MOVL C00866 V=7.0 ACC=20 DEC=20
MOVL C00867 V=7.0 ACC=20 DEC=20
MOVL C00868 V=7.0 ACC=20 DEC=20
MOVL C00869 V=7.0 ACC=20 DEC=20
MOVL C00870 V=7.0 ACC=20 DEC=20
MOVL C00871 V=7.0 ACC=20 DEC=20
MOVL C00872 V=7.0 ACC=20 DEC=20
MOVL C00873 V=7.0 ACC=20 DEC=20
MOVL C00874 V=7.0 ACC=20 DEC=20
MOVL C00875 V=7.0 ACC=20 DEC=20
MOVL C00876 V=7.0 ACC=20 DEC=20
MOVL C00877 V=7.0 ACC=20 DEC=20
MOVL C00878 V=7.0 PL=1
MOVL C00879 V=7.0 ACC=20 DEC=20
MOVL C00880 V=7.0 ACC=20 DEC=20
MOVL C00881 V=7.0 ACC=20 DEC=20
MOVL C00882 V=7.0 ACC=20 DEC=20
MOVL C00883 V=7.0 ACC=20 DEC=20
MOVL C00884 V=7.0 ACC=20 DEC=20
MOVL C00885 V=7.0 ACC=20 DEC=20
MOVL C00886 V=7.0 ACC=20 DEC=20
MOVL C00887 V=7.0 ACC=20 DEC=20
MOVL C00888 V=11.0 ACC=20 DEC=20
MOVC C00889 V=11.0 ACC=20 DEC=20
MOVC C00890 V=11.0 ACC=20 DEC=20
MOVC C00891 V=11.0 ACC=20 DEC=20
MOVL C00892 V=7.0 ACC=20 DEC=20
MOVL C00893 V=7.0 ACC=20 DEC=20
MOVL C00894 V=7.0 ACC=20 DEC=20
MOVL C00895 V=7.0 ACC=20 DEC=20
MOVL C00896 V=7.0 ACC=20 DEC=20
MOVL C00897 V=7.0 ACC=20 DEC=20
MOVL C00898 V=7.0 ACC=20 DEC=20
MOVL C00899 V=7.0 ACC=20 DEC=20
MOVL C00900 V=7.0 ACC=20 DEC=20
MOVL C00901 V=7.0 ACC=20 DEC=20
MOVL C00902 V=7.0 ACC=20 DEC=20
MOVL C00903 V=7.0 ACC=20 DEC=20
MOVL C00904 V=7.0 ACC=20 DEC=20
MOVL C00905 V=7.0 ACC=20 DEC=20
MOVL C00906 V=7.0 ACC=20 DEC=20
MOVL C00907 V=7.0 ACC=20 DEC=20
MOVL C00908 V=7.0 ACC=20 DEC=20
MOVL C00909 V=7.0 ACC=20 DEC=20
MOVL C00910 V=7.0 ACC=20 DEC=20
MOVL C00911 V=7.0 ACC=20 DEC=20
ARCOF
TIMER T=30.00
MOVL C00912 V=11.0 ACC=20 DEC=20
*LAG11
MACRO1 MJ#(0) ARGF2
ARCON
MOVL C00913 V=7.0 ACC=20 DEC=20
MOVL C00914 V=7.0 ACC=20 DEC=20
MOVL C00915 V=7.0 ACC=20 DEC=20
MOVL C00916 V=7.0 ACC=20 DEC=20
MOVL C00917 V=7.0 ACC=20 DEC=20
MOVL C00918 V=7.0 ACC=20 DEC=20
MOVL C00919 V=7.0 ACC=20 DEC=20
MOVL C00920 V=7.0 ACC=20 DEC=20
MOVL C00921 V=7.0 ACC=20 DEC=20
MOVL C00922 V=7.0 ACC=20 DEC=20
MOVL C00923 V=7.0 ACC=20 DEC=20
MOVL C00924 V=7.0 ACC=20 DEC=20
MOVL C00925 V=7.0 ACC=20 DEC=20
MOVL C00926 V=7.0 ACC=20 DEC=20
MOVL C00927 V=7.0 ACC=20 DEC=20
MOVL C00928 V=7.0 ACC=20 DEC=20
MOVL C00929 V=7.0 ACC=20 DEC=20
MOVL C00930 V=7.0 ACC=20 DEC=20
MOVL C00931 V=7.0 ACC=20 DEC=20
MOVL C00932 V=11.0 ACC=20 DEC=20
MOVC C00933 V=11.0 ACC=20 DEC=20
MOVC C00934 V=11.0 ACC=20 DEC=20
MOVC C00935 V=11.0 ACC=20 DEC=20
MOVL C00936 V=7.0 ACC=20 DEC=20
MOVL C00937 V=7.0 ACC=20 DEC=20
MOVL C00938 V=7.0 ACC=20 DEC=20
MOVL C00939 V=7.0 ACC=20 DEC=20
MOVL C00940 V=7.0 ACC=20 DEC=20
MOVL C00941 V=7.0 ACC=20 DEC=20
MOVL C00942 V=7.0 ACC=20 DEC=20
MOVL C00943 V=7.0 ACC=20 DEC=20
MOVL C00944 V=7.0 ACC=20 DEC=20
MOVL C00945 V=7.0 PL=1
MOVL C00946 V=7.0 ACC=20 DEC=20
MOVL C00947 V=7.0 ACC=20 DEC=20
MOVL C00948 V=7.0 ACC=20 DEC=20
MOVL C00949 V=7.0 ACC=20 DEC=20
MOVL C00950 V=7.0 ACC=20 DEC=20
MOVL C00951 V=7.0 ACC=20 DEC=20
MOVL C00952 V=7.0 ACC=20 DEC=20
MOVL C00953 V=7.0 ACC=20 DEC=20
MOVL C00954 V=7.0 ACC=20 DEC=20
MOVL C00955 V=7.0 ACC=20 DEC=20
MOVL C00956 V=7.0 ACC=20 DEC=20
MOVL C00957 V=7.0 ACC=20 DEC=20
MOVL C00958 V=7.0 ACC=20 DEC=20
MOVL C00959 V=7.0 ACC=20 DEC=20
MOVL C00960 V=7.0 ACC=20 DEC=20
MOVL C00961 V=7.0 ACC=20 DEC=20
MOVL C00962 V=7.0 ACC=20 DEC=20
MOVL C00963 V=7.0 ACC=20 DEC=20
MOVL C00964 V=7.0 ACC=20 DEC=20
MOVL C00965 V=7.0 ACC=20 DEC=20
MOVL C00966 V=7.0 ACC=20 DEC=20
MOVL C00967 V=11.0 ACC=20 DEC=20
MOVC C00968 V=11.0 ACC=20 DEC=20
MOVC C00969 V=11.0 ACC=20 DEC=20
MOVC C00970 V=11.0 ACC=20 DEC=20
MOVL C00971 V=7.0 ACC=20 DEC=20
MOVL C00972 V=7.0 ACC=20 DEC=20
MOVL C00973 V=7.0 ACC=20 DEC=20
MOVL C00974 V=7.0 ACC=20 DEC=20
MOVL C00975 V=7.0 ACC=20 DEC=20
MOVL C00976 V=7.0 ACC=20 DEC=20
MOVL C00977 V=7.0 ACC=20 DEC=20
MOVL C00978 V=7.0 ACC=20 DEC=20
MOVL C00979 V=7.0 ACC=20 DEC=20
MOVL C00980 V=7.0 ACC=20 DEC=20
MOVL C00981 V=7.0 ACC=20 DEC=20
MOVL C00982 V=7.0 ACC=20 DEC=20
MOVL C00983 V=7.0 ACC=20 DEC=20
MOVL C00984 V=7.0 ACC=20 DEC=20
MOVL C00985 V=7.0 ACC=20 DEC=20
MOVL C00986 V=7.0 ACC=20 DEC=20
MOVL C00987 V=7.0 ACC=20 DEC=20
MOVL C00988 V=7.0 ACC=20 DEC=20
MOVL C00989 V=7.0 ACC=20 DEC=20
MOVL C00990 V=7.0 ACC=20 DEC=20
MOVL C00991 V=7.0 ACC=20 DEC=20
MOVL C00992 V=7.0 PL=1
MOVL C00993 V=7.0 ACC=20 DEC=20
MOVL C00994 V=7.0 ACC=20 DEC=20
MOVL C00995 V=7.0 ACC=20 DEC=20
MOVL C00996 V=7.0 ACC=20 DEC=20
MOVL C00997 V=7.0 ACC=20 DEC=20
MOVL C00998 V=7.0 ACC=20 DEC=20
MOVL C00999 V=7.0 ACC=20 DEC=20
MOVL C01000 V=7.0 ACC=20 DEC=20
MOVL C01001 V=7.0 ACC=20 DEC=20
MOVL C01002 V=7.0 ACC=20 DEC=20
ARCOF
TIMER T=30.00
MOVL C01003 V=11.0 ACC=20 DEC=20
*LAG12
MACRO1 MJ#(0) ARGF2
ARCON
MOVL C01004 V=7.0 ACC=20 DEC=20
MOVL C01005 V=7.0 ACC=20 DEC=20
MOVL C01006 V=7.0 ACC=20 DEC=20
MOVL C01007 V=7.0 ACC=20 DEC=20
MOVL C01008 V=7.0 ACC=20 DEC=20
MOVL C01009 V=7.0 ACC=20 DEC=20
MOVL C01010 V=7.0 ACC=20 DEC=20
MOVL C01011 V=7.0 ACC=20 DEC=20
MOVL C01012 V=7.0 ACC=20 DEC=20
MOVL C01013 V=7.0 PL=1
MOVL C01014 V=7.0 ACC=20 DEC=20
MOVL C01015 V=7.0 ACC=20 DEC=20
MOVL C01016 V=7.0 ACC=20 DEC=20
MOVL C01017 V=7.0 ACC=20 DEC=20
MOVL C01018 V=7.0 ACC=20 DEC=20
MOVL C01019 V=7.0 ACC=20 DEC=20
MOVL C01020 V=7.0 ACC=20 DEC=20
MOVL C01021 V=7.0 ACC=20 DEC=20
MOVL C01022 V=7.0 ACC=20 DEC=20
MOVL C01023 V=7.0 ACC=20 DEC=20
MOVL C01024 V=7.0 ACC=20 DEC=20
MOVL C01025 V=7.0 ACC=20 DEC=20
MOVL C01026 V=7.0 ACC=20 DEC=20
MOVL C01027 V=7.0 ACC=20 DEC=20
MOVL C01028 V=7.0 ACC=20 DEC=20
MOVL C01029 V=7.0 ACC=20 DEC=20
MOVL C01030 V=7.0 ACC=20 DEC=20
MOVL C01031 V=7.0 ACC=20 DEC=20
MOVL C01032 V=7.0 ACC=20 DEC=20
MOVL C01033 V=7.0 ACC=20 DEC=20
MOVL C01034 V=7.0 ACC=20 DEC=20
MOVL C01035 V=11.0 ACC=20 DEC=20
MOVC C01036 V=11.0 ACC=20 DEC=20
MOVC C01037 V=11.0 ACC=20 DEC=20
MOVC C01038 V=11.0 ACC=20 DEC=20
MOVL C01039 V=7.0 ACC=20 DEC=20
MOVL C01040 V=7.0 ACC=20 DEC=20
MOVL C01041 V=7.0 ACC=20 DEC=20
MOVL C01042 V=7.0 ACC=20 DEC=20
MOVL C01043 V=7.0 ACC=20 DEC=20
MOVL C01044 V=7.0 ACC=20 DEC=20
MOVL C01045 V=7.0 ACC=20 DEC=20
MOVL C01046 V=7.0 ACC=20 DEC=20
MOVL C01047 V=7.0 ACC=20 DEC=20
MOVL C01048 V=7.0 ACC=20 DEC=20
MOVL C01049 V=7.0 ACC=20 DEC=20
MOVL C01050 V=7.0 ACC=20 DEC=20
MOVL C01051 V=7.0 ACC=20 DEC=20
MOVL C01052 V=7.0 ACC=20 DEC=20
MOVL C01053 V=7.0 ACC=20 DEC=20
MOVL C01054 V=7.0 ACC=20 DEC=20
MOVL C01055 V=7.0 ACC=20 DEC=20
MOVL C01056 V=7.0 ACC=20 DEC=20
MOVL C01057 V=7.0 ACC=20 DEC=20
MOVL C01058 V=7.0 ACC=20 DEC=20
MOVL C01059 V=7.0 ACC=20 DEC=20
MOVL C01060 V=7.0 PL=1
MOVL C01061 V=7.0 ACC=20 DEC=20
MOVL C01062 V=7.0 ACC=20 DEC=20
MOVL C01063 V=7.0 ACC=20 DEC=20
MOVL C01064 V=7.0 ACC=20 DEC=20
MOVL C01065 V=7.0 ACC=20 DEC=20
MOVL C01066 V=7.0 ACC=20 DEC=20
MOVL C01067 V=7.0 ACC=20 DEC=20
MOVL C01068 V=7.0 ACC=20 DEC=20
MOVL C01069 V=7.0 ACC=20 DEC=20
MOVL C01070 V=11.0 ACC=20 DEC=20
MOVC C01071 V=11.0 ACC=20 DEC=20
MOVC C01072 V=11.0 ACC=20 DEC=20
MOVC C01073 V=11.0 ACC=20 DEC=20
MOVL C01074 V=7.0 ACC=20 DEC=20
MOVL C01075 V=7.0 ACC=20 DEC=20
MOVL C01076 V=7.0 ACC=20 DEC=20
MOVL C01077 V=7.0 ACC=20 DEC=20
MOVL C01078 V=7.0 ACC=20 DEC=20
MOVL C01079 V=7.0 ACC=20 DEC=20
MOVL C01080 V=7.0 ACC=20 DEC=20
MOVL C01081 V=7.0 ACC=20 DEC=20
MOVL C01082 V=7.0 ACC=20 DEC=20
MOVL C01083 V=7.0 ACC=20 DEC=20
MOVL C01084 V=7.0 ACC=20 DEC=20
MOVL C01085 V=7.0 ACC=20 DEC=20
MOVL C01086 V=7.0 ACC=20 DEC=20
MOVL C01087 V=7.0 ACC=20 DEC=20
MOVL C01088 V=7.0 ACC=20 DEC=20
MOVL C01089 V=7.0 ACC=20 DEC=20
MOVL C01090 V=7.0 ACC=20 DEC=20
MOVL C01091 V=7.0 ACC=20 DEC=20
MOVL C01092 V=7.0 ACC=20 DEC=20
MOVL C01093 V=7.0 ACC=20 DEC=20
ARCOF
TIMER T=30.00
MOVL C01094 V=11.0 ACC=20 DEC=20
*LAG13
MACRO1 MJ#(0) ARGF2
ARCON
MOVL C01095 V=7.0 ACC=20 DEC=20
MOVL C01096 V=7.0 ACC=20 DEC=20
MOVL C01097 V=7.0 ACC=20 DEC=20
MOVL C01098 V=7.0 ACC=20 DEC=20
MOVL C01099 V=7.0 ACC=20 DEC=20
MOVL C01100 V=7.0 ACC=20 DEC=20
MOVL C01101 V=7.0 ACC=20 DEC=20
MOVL C01102 V=7.0 ACC=20 DEC=20
MOVL C01103 V=7.0 ACC=20 DEC=20
MOVL C01104 V=7.0 ACC=20 DEC=20
MOVL C01105 V=7.0 ACC=20 DEC=20
MOVL C01106 V=7.0 ACC=20 DEC=20
MOVL C01107 V=7.0 ACC=20 DEC=20
MOVL C01108 V=7.0 ACC=20 DEC=20
MOVL C01109 V=7.0 ACC=20 DEC=20
MOVL C01110 V=7.0 ACC=20 DEC=20
MOVL C01111 V=7.0 ACC=20 DEC=20
MOVL C01112 V=7.0 ACC=20 DEC=20
MOVL C01113 V=7.0 ACC=20 DEC=20
MOVL C01114 V=11.0 ACC=20 DEC=20
MOVC C01115 V=11.0 ACC=20 DEC=20
MOVC C01116 V=11.0 ACC=20 DEC=20
MOVC C01117 V=11.0 ACC=20 DEC=20
MOVL C01118 V=7.0 ACC=20 DEC=20
MOVL C01119 V=7.0 ACC=20 DEC=20
MOVL C01120 V=7.0 ACC=20 DEC=20
MOVL C01121 V=7.0 ACC=20 DEC=20
MOVL C01122 V=7.0 ACC=20 DEC=20
MOVL C01123 V=7.0 ACC=20 DEC=20
MOVL C01124 V=7.0 ACC=20 DEC=20
MOVL C01125 V=7.0 ACC=20 DEC=20
MOVL C01126 V=7.0 ACC=20 DEC=20
MOVL C01127 V=7.0 PL=1
MOVL C01128 V=7.0 ACC=20 DEC=20
MOVL C01129 V=7.0 ACC=20 DEC=20
MOVL C01130 V=7.0 ACC=20 DEC=20
MOVL C01131 V=7.0 ACC=20 DEC=20
MOVL C01132 V=7.0 ACC=20 DEC=20
MOVL C01133 V=7.0 ACC=20 DEC=20
MOVL C01134 V=7.0 ACC=20 DEC=20
MOVL C01135 V=7.0 ACC=20 DEC=20
MOVL C01136 V=7.0 ACC=20 DEC=20
MOVL C01137 V=7.0 ACC=20 DEC=20
MOVL C01138 V=7.0 ACC=20 DEC=20
MOVL C01139 V=7.0 ACC=20 DEC=20
MOVL C01140 V=7.0 ACC=20 DEC=20
MOVL C01141 V=7.0 ACC=20 DEC=20
MOVL C01142 V=7.0 ACC=20 DEC=20
MOVL C01143 V=7.0 ACC=20 DEC=20
MOVL C01144 V=7.0 ACC=20 DEC=20
MOVL C01145 V=7.0 ACC=20 DEC=20
MOVL C01146 V=7.0 ACC=20 DEC=20
MOVL C01147 V=7.0 ACC=20 DEC=20
MOVL C01148 V=7.0 ACC=20 DEC=20
MOVL C01149 V=11.0 ACC=20 DEC=20
MOVC C01150 V=11.0 ACC=20 DEC=20
MOVC C01151 V=11.0 ACC=20 DEC=20
MOVC C01152 V=11.0 ACC=20 DEC=20
MOVL C01153 V=7.0 ACC=20 DEC=20
MOVL C01154 V=7.0 ACC=20 DEC=20
MOVL C01155 V=7.0 ACC=20 DEC=20
MOVL C01156 V=7.0 ACC=20 DEC=20
MOVL C01157 V=7.0 ACC=20 DEC=20
MOVL C01158 V=7.0 ACC=20 DEC=20
MOVL C01159 V=7.0 ACC=20 DEC=20
MOVL C01160 V=7.0 ACC=20 DEC=20
MOVL C01161 V=7.0 ACC=20 DEC=20
MOVL C01162 V=7.0 ACC=20 DEC=20
MOVL C01163 V=7.0 ACC=20 DEC=20
MOVL C01164 V=7.0 ACC=20 DEC=20
MOVL C01165 V=7.0 ACC=20 DEC=20
MOVL C01166 V=7.0 ACC=20 DEC=20
MOVL C01167 V=7.0 ACC=20 DEC=20
MOVL C01168 V=7.0 ACC=20 DEC=20
MOVL C01169 V=7.0 ACC=20 DEC=20
MOVL C01170 V=7.0 ACC=20 DEC=20
MOVL C01171 V=7.0 ACC=20 DEC=20
MOVL C01172 V=7.0 ACC=20 DEC=20
MOVL C01173 V=7.0 ACC=20 DEC=20
MOVL C01174 V=7.0 PL=1
MOVL C01175 V=7.0 ACC=20 DEC=20
MOVL C01176 V=7.0 ACC=20 DEC=20
MOVL C01177 V=7.0 ACC=20 DEC=20
MOVL C01178 V=7.0 ACC=20 DEC=20
MOVL C01179 V=7.0 ACC=20 DEC=20
MOVL C01180 V=7.0 ACC=20 DEC=20
MOVL C01181 V=7.0 ACC=20 DEC=20
MOVL C01182 V=7.0 ACC=20 DEC=20
MOVL C01183 V=7.0 ACC=20 DEC=20
MOVL C01184 V=7.0 ACC=20 DEC=20
ARCOF
TIMER T=30.00
MOVL C01185 V=11.0 ACC=20 DEC=20
*LAG14
MACRO1 MJ#(0) ARGF2
ARCON
MOVL C01186 V=7.0 ACC=20 DEC=20
MOVL C01187 V=7.0 ACC=20 DEC=20
MOVL C01188 V=7.0 ACC=20 DEC=20
MOVL C01189 V=7.0 ACC=20 DEC=20
MOVL C01190 V=7.0 ACC=20 DEC=20
MOVL C01191 V=7.0 ACC=20 DEC=20
MOVL C01192 V=7.0 ACC=20 DEC=20
MOVL C01193 V=7.0 ACC=20 DEC=20
MOVL C01194 V=7.0 ACC=20 DEC=20
MOVL C01195 V=7.0 PL=1
MOVL C01196 V=7.0 ACC=20 DEC=20
MOVL C01197 V=7.0 ACC=20 DEC=20
MOVL C01198 V=7.0 ACC=20 DEC=20
MOVL C01199 V=7.0 ACC=20 DEC=20
MOVL C01200 V=7.0 ACC=20 DEC=20
MOVL C01201 V=7.0 ACC=20 DEC=20
MOVL C01202 V=7.0 ACC=20 DEC=20
MOVL C01203 V=7.0 ACC=20 DEC=20
MOVL C01204 V=7.0 ACC=20 DEC=20
MOVL C01205 V=7.0 ACC=20 DEC=20
MOVL C01206 V=7.0 ACC=20 DEC=20
MOVL C01207 V=7.0 ACC=20 DEC=20
MOVL C01208 V=7.0 ACC=20 DEC=20
MOVL C01209 V=7.0 ACC=20 DEC=20
MOVL C01210 V=7.0 ACC=20 DEC=20
MOVL C01211 V=7.0 ACC=20 DEC=20
MOVL C01212 V=7.0 ACC=20 DEC=20
MOVL C01213 V=7.0 ACC=20 DEC=20
MOVL C01214 V=7.0 ACC=20 DEC=20
MOVL C01215 V=7.0 ACC=20 DEC=20
MOVL C01216 V=7.0 ACC=20 DEC=20
MOVL C01217 V=11.0 ACC=20 DEC=20
MOVC C01218 V=11.0 ACC=20 DEC=20
MOVC C01219 V=11.0 ACC=20 DEC=20
MOVC C01220 V=11.0 ACC=20 DEC=20
MOVL C01221 V=7.0 ACC=20 DEC=20
MOVL C01222 V=7.0 ACC=20 DEC=20
MOVL C01223 V=7.0 ACC=20 DEC=20
MOVL C01224 V=7.0 ACC=20 DEC=20
MOVL C01225 V=7.0 ACC=20 DEC=20
MOVL C01226 V=7.0 ACC=20 DEC=20
MOVL C01227 V=7.0 ACC=20 DEC=20
MOVL C01228 V=7.0 ACC=20 DEC=20
MOVL C01229 V=7.0 ACC=20 DEC=20
MOVL C01230 V=7.0 ACC=20 DEC=20
MOVL C01231 V=7.0 ACC=20 DEC=20
MOVL C01232 V=7.0 ACC=20 DEC=20
MOVL C01233 V=7.0 ACC=20 DEC=20
MOVL C01234 V=7.0 ACC=20 DEC=20
MOVL C01235 V=7.0 ACC=20 DEC=20
MOVL C01236 V=7.0 ACC=20 DEC=20
MOVL C01237 V=7.0 ACC=20 DEC=20
MOVL C01238 V=7.0 ACC=20 DEC=20
MOVL C01239 V=7.0 ACC=20 DEC=20
MOVL C01240 V=7.0 ACC=20 DEC=20
MOVL C01241 V=7.0 ACC=20 DEC=20
MOVL C01242 V=7.0 PL=1
MOVL C01243 V=7.0 ACC=20 DEC=20
MOVL C01244 V=7.0 ACC=20 DEC=20
MOVL C01245 V=7.0 ACC=20 DEC=20
MOVL C01246 V=7.0 ACC=20 DEC=20
MOVL C01247 V=7.0 ACC=20 DEC=20
MOVL C01248 V=7.0 ACC=20 DEC=20
MOVL C01249 V=7.0 ACC=20 DEC=20
MOVL C01250 V=7.0 ACC=20 DEC=20
MOVL C01251 V=7.0 ACC=20 DEC=20
MOVL C01252 V=11.0 ACC=20 DEC=20
MOVC C01253 V=11.0 ACC=20 DEC=20
MOVC C01254 V=11.0 ACC=20 DEC=20
MOVC C01255 V=11.0 ACC=20 DEC=20
MOVL C01256 V=7.0 ACC=20 DEC=20
MOVL C01257 V=7.0 ACC=20 DEC=20
MOVL C01258 V=7.0 ACC=20 DEC=20
MOVL C01259 V=7.0 ACC=20 DEC=20
MOVL C01260 V=7.0 ACC=20 DEC=20
MOVL C01261 V=7.0 ACC=20 DEC=20
MOVL C01262 V=7.0 ACC=20 DEC=20
MOVL C01263 V=7.0 ACC=20 DEC=20
MOVL C01264 V=7.0 ACC=20 DEC=20
MOVL C01265 V=7.0 ACC=20 DEC=20
MOVL C01266 V=7.0 ACC=20 DEC=20
MOVL C01267 V=7.0 ACC=20 DEC=20
MOVL C01268 V=7.0 ACC=20 DEC=20
MOVL C01269 V=7.0 ACC=20 DEC=20
MOVL C01270 V=7.0 ACC=20 DEC=20
MOVL C01271 V=7.0 ACC=20 DEC=20
MOVL C01272 V=7.0 ACC=20 DEC=20
MOVL C01273 V=7.0 ACC=20 DEC=20
MOVL C01274 V=7.0 ACC=20 DEC=20
MOVL C01275 V=7.0 ACC=20 DEC=20
ARCOF
TIMER T=30.00
MOVL C01276 V=11.0 ACC=20 DEC=20
*LAG15
MACRO1 MJ#(0) ARGF2
ARCON
MOVL C01277 V=7.0 ACC=20 DEC=20
MOVL C01278 V=7.0 ACC=20 DEC=20
MOVL C01279 V=7.0 ACC=20 DEC=20
MOVL C01280 V=7.0 ACC=20 DEC=20
MOVL C01281 V=7.0 ACC=20 DEC=20
MOVL C01282 V=7.0 ACC=20 DEC=20
MOVL C01283 V=7.0 ACC=20 DEC=20
MOVL C01284 V=7.0 ACC=20 DEC=20
MOVL C01285 V=7.0 ACC=20 DEC=20
MOVL C01286 V=7.0 ACC=20 DEC=20
MOVL C01287 V=7.0 ACC=20 DEC=20
MOVL C01288 V=7.0 ACC=20 DEC=20
MOVL C01289 V=7.0 ACC=20 DEC=20
MOVL C01290 V=7.0 ACC=20 DEC=20
MOVL C01291 V=7.0 ACC=20 DEC=20
MOVL C01292 V=7.0 ACC=20 DEC=20
MOVL C01293 V=7.0 ACC=20 DEC=20
MOVL C01294 V=7.0 ACC=20 DEC=20
MOVL C01295 V=7.0 ACC=20 DEC=20
MOVL C01296 V=11.0 ACC=20 DEC=20
MOVC C01297 V=11.0 ACC=20 DEC=20
MOVC C01298 V=11.0 ACC=20 DEC=20
MOVC C01299 V=11.0 ACC=20 DEC=20
MOVL C01300 V=7.0 ACC=20 DEC=20
MOVL C01301 V=7.0 ACC=20 DEC=20
MOVL C01302 V=7.0 ACC=20 DEC=20
MOVL C01303 V=7.0 ACC=20 DEC=20
MOVL C01304 V=7.0 ACC=20 DEC=20
MOVL C01305 V=7.0 ACC=20 DEC=20
MOVL C01306 V=7.0 ACC=20 DEC=20
MOVL C01307 V=7.0 ACC=20 DEC=20
MOVL C01308 V=7.0 ACC=20 DEC=20
MOVL C01309 V=7.0 PL=1
MOVL C01310 V=7.0 ACC=20 DEC=20
MOVL C01311 V=7.0 ACC=20 DEC=20
MOVL C01312 V=7.0 ACC=20 DEC=20
MOVL C01313 V=7.0 ACC=20 DEC=20
MOVL C01314 V=7.0 ACC=20 DEC=20
MOVL C01315 V=7.0 ACC=20 DEC=20
MOVL C01316 V=7.0 ACC=20 DEC=20
MOVL C01317 V=7.0 ACC=20 DEC=20
MOVL C01318 V=7.0 ACC=20 DEC=20
MOVL C01319 V=7.0 ACC=20 DEC=20
MOVL C01320 V=7.0 ACC=20 DEC=20
MOVL C01321 V=7.0 ACC=20 DEC=20
MOVL C01322 V=7.0 ACC=20 DEC=20
MOVL C01323 V=7.0 ACC=20 DEC=20
MOVL C01324 V=7.0 ACC=20 DEC=20
MOVL C01325 V=7.0 ACC=20 DEC=20
MOVL C01326 V=7.0 ACC=20 DEC=20
MOVL C01327 V=7.0 ACC=20 DEC=20
MOVL C01328 V=7.0 ACC=20 DEC=20
MOVL C01329 V=7.0 ACC=20 DEC=20
MOVL C01330 V=7.0 ACC=20 DEC=20
MOVL C01331 V=11.0 ACC=20 DEC=20
MOVC C01332 V=11.0 ACC=20 DEC=20
MOVC C01333 V=11.0 ACC=20 DEC=20
MOVC C01334 V=11.0 ACC=20 DEC=20
MOVL C01335 V=7.0 ACC=20 DEC=20
MOVL C01336 V=7.0 ACC=20 DEC=20
MOVL C01337 V=7.0 ACC=20 DEC=20
MOVL C01338 V=7.0 ACC=20 DEC=20
MOVL C01339 V=7.0 ACC=20 DEC=20
MOVL C01340 V=7.0 ACC=20 DEC=20
MOVL C01341 V=7.0 ACC=20 DEC=20
MOVL C01342 V=7.0 ACC=20 DEC=20
MOVL C01343 V=7.0 ACC=20 DEC=20
MOVL C01344 V=7.0 ACC=20 DEC=20
MOVL C01345 V=7.0 ACC=20 DEC=20
MOVL C01346 V=7.0 ACC=20 DEC=20
MOVL C01347 V=7.0 ACC=20 DEC=20
MOVL C01348 V=7.0 ACC=20 DEC=20
MOVL C01349 V=7.0 ACC=20 DEC=20
MOVL C01350 V=7.0 ACC=20 DEC=20
MOVL C01351 V=7.0 ACC=20 DEC=20
MOVL C01352 V=7.0 ACC=20 DEC=20
MOVL C01353 V=7.0 ACC=20 DEC=20
MOVL C01354 V=7.0 ACC=20 DEC=20
MOVL C01355 V=7.0 ACC=20 DEC=20
MOVL C01356 V=7.0 PL=1
MOVL C01357 V=7.0 ACC=20 DEC=20
MOVL C01358 V=7.0 ACC=20 DEC=20
MOVL C01359 V=7.0 ACC=20 DEC=20
MOVL C01360 V=7.0 ACC=20 DEC=20
MOVL C01361 V=7.0 ACC=20 DEC=20
MOVL C01362 V=7.0 ACC=20 DEC=20
MOVL C01363 V=7.0 ACC=20 DEC=20
MOVL C01364 V=7.0 ACC=20 DEC=20
MOVL C01365 V=7.0 ACC=20 DEC=20
MOVL C01366 V=7.0 ACC=20 DEC=20
ARCOF
TIMER T=30.00
MOVL C01367 V=11.0 ACC=20 DEC=20
MOVJ C01368 VJ=0.78
END
